GLOBALCONSTANTS SubStrings (* Global constants *)
  (* Standard: 61499-1 *)
  (* Version 1.0, 2026-11-04, Franz Höpfinger, Meisterschulen am Ostbahnhof *)
  PACKAGE Meins::Servo_AI4_Calibrate_OPC;
  VAR_GLOBAL CONSTANT
    SAI4_RAW_WRITE : WSTRING := "opc_ua[WRITE;/Objects/ServoAI4/RAW,1:s=SAI4_RAW]"; (* Rohwert AI4 0-4095 *)
    SAI4_CAL_WRITE : WSTRING := "opc_ua[WRITE;/Objects/ServoAI4/CAL,1:s=SAI4_CAL]"; (* kalibrierter Wert AI4 = Sollwinkel *)
    SAI4_MIN_METHOD : WSTRING := "opc_ua[CREATE_METHOD;/Objects/ServoAI4/MINMethod,1:s=SAI4_MIN_METHOD]"; (* Trigger C_MIN *)
    SAI4_MID_METHOD : WSTRING := "opc_ua[CREATE_METHOD;/Objects/ServoAI4/MIDMethod,1:s=SAI4_MID_METHOD]"; (* Trigger C_MID *)
    SAI4_MAX_METHOD : WSTRING := "opc_ua[CREATE_METHOD;/Objects/ServoAI4/MAXMethod,1:s=SAI4_MAX_METHOD]"; (* Trigger C_MAX *)
    SAI4_MINREF_READ : WSTRING := "opc_ua[READ;/Objects/ServoAI4/MINREFExt,1:s=SAI4_MINREF_EXT]"; (* MIN_REF vom Dashboard *)
    SAI4_MINREF_WRITE : WSTRING := "opc_ua[WRITE;/Objects/ServoAI4/MINREF,1:s=SAI4_MINREF]"; (* MIN_REF Echo *)
    SAI4_MIDREF_READ : WSTRING := "opc_ua[READ;/Objects/ServoAI4/MIDREFExt,1:s=SAI4_MIDREF_EXT]"; (* MID_REF vom Dashboard *)
    SAI4_MIDREF_WRITE : WSTRING := "opc_ua[WRITE;/Objects/ServoAI4/MIDREF,1:s=SAI4_MIDREF]"; (* MID_REF Echo *)
    SAI4_MAXREF_READ : WSTRING := "opc_ua[READ;/Objects/ServoAI4/MAXREFExt,1:s=SAI4_MAXREF_EXT]"; (* MAX_REF vom Dashboard *)
    SAI4_MAXREF_WRITE : WSTRING := "opc_ua[WRITE;/Objects/ServoAI4/MAXREF,1:s=SAI4_MAXREF]"; (* MAX_REF Echo *)
    SAI4_MIN_RAW_WRITE : WSTRING := "opc_ua[WRITE;/Objects/ServoAI4/MINRAW,1:s=SAI4_MIN_RAW]"; (* Rohwert am MIN-Punkt *)
    SAI4_MID_RAW_WRITE : WSTRING := "opc_ua[WRITE;/Objects/ServoAI4/MIDRAW,1:s=SAI4_MID_RAW]"; (* Rohwert am MID-Punkt *)
    SAI4_MAX_RAW_WRITE : WSTRING := "opc_ua[WRITE;/Objects/ServoAI4/MAXRAW,1:s=SAI4_MAX_RAW]"; (* Rohwert am MAX-Punkt *)
    SAI4_ANGLE : WSTRING := "opc_ua[WRITE;/Objects/ServoAI4/ANGLE,1:s=SAI4_ANGLE]"; (* angewendeter Winkel Q2 (Echo) *)
  END_VAR
END_GLOBALCONSTANTS
